Omron Sysmac Studio project medina sin node con todo (Sysmac Studio 1.64.0.64008, StandardProject)

# Controller new_Controller_0: NX102-1020 version 1.60
Axis MC_Axis000, settings changed from default: AxisType=ServoType, FunctionLimit=SingleAxisPTP, UnitsConversion=EnumElement5, UnitsNumerator=8388608, ReducerUse=EnumElement2, TravelDistancePerWorkRotation=180, WorkGearRatio=100, MotorGearRatio=198, MaxVelocity=20, MaxJogVelocity=20, CountMode=EnumElement2, ModuloMAXPosition=360, ModuloMINPosition=0, EncoderTypes=Abs
Axis MC_Axis001, settings changed from default: AxisNumber=1, AxisType=ServoType, FunctionLimit=SingleAxisPTP, UnitsConversion=EnumElement2, UnitsNumerator=8388608, UnitsDenominator=290, MaxVelocity=10, MaxJogVelocity=10, EncoderTypes=Abs
Task PrimaryTask (priority 4, period or condition 2000): Programa0, main
Task PeriodicTask0 (priority 17, period or condition 20000): AMR
Library TMEthernetIP_v2.0.0 2.0.0 (contents left out)
Library ARCL_Comms_Lib 1.3.0 (contents left out)

TYPE RfidCommand : STRUCT
    CommExec : WORD;
    CmdCode : WORD;
    CmdParam1 : WORD;
    CmdParam2 : WORD;
    CmdData : array[0..15] of word;
END_STRUCT END_TYPE
TYPE RfidResponse : STRUCT
    RfidStatus : WORD;
    RfidErrorCode : WORD;
    RfidRespInfo1 : WORD;
    RfidRespInfo2 : WORD;
    RfidRespData : array[0..15] of WORD;
END_STRUCT END_TYPE
TYPE RFID_Status : UNION
    Status_reg : word;
    Status_bits : ARRAY[0..15] OF BOOL;
END_UNION END_TYPE
TYPE CmdRFID : (Read_ID := 1, Read_data := 2, Write_Data := 3, LockRfid := 4, Data_fill := 5, Overwrite_control := 6, Restore_data := 7, Copy_data := 8, Initialize := 4096, Set_RF_Comm_Settings := 4097, Get_RF_tag_comm := 4098, Set_multi_Reades := 4099, Get_multi_reader := 4100, Get_model_information := 8192, Get_firmware_version := 8193, Get_operating_time := 8194, Measure_noise := 8195, Get_comd_error_log := 8196, Get_restore_infomation := 8197, Get_multireader_status := 8198, Reset := 12288); END_TYPE
TYPE Status_struct : STRUCT
    Datos_bits : ARRAY[0..15] OF BOOL;
END_STRUCT END_TYPE
TYPE stCarouselSlot : STRUCT
    RoomID : INT;
    MedID : INT;
    IsLoaded : BOOL;
    IsDelivered : BOOL;
END_STRUCT END_TYPE

VAR_GLOBAL
    DataFromRFID : RfidResponse;  (* network input *)
    ArrayFromTM : array[0..491] of byte;  (* network input *)
    ArrayToTM : array[0..295] of byte;  (* network output *)
    StructFromTM : ATC_E\TMEthernetIP\FromTM;
    StructToTM : ATC_E\TMEthernetIP\ToTM;
    DataToRFID : RfidCommand;  (* network output *)
END_VAR
VAR_GLOBAL CONSTANT
    MC_Axis000 : _sAXIS_REF;  (* at MC://_MC_AX[0] *)
    MC_Axis001 : _sAXIS_REF;  (* at MC://_MC_AX[1] *)
END_VAR
VAR_GLOBAL
    habitaciones : ARRAY[0..9] OF int;  (* network output *)
    medicamentos : ARRAY[0..9] OF int;  (* network output *)
    test_escritura : INT;  (* published *)
    Carrusel : ARRAY[0..9] OF stCarouselSlot;
    etapa : INT;
    activar : BOOL;
    done_amr : BOOL;
    pos_carrusel : LREAL;
    pos_trampilla : LREAL;
    done_carrusel : BOOL;
    done_trampilla : BOOL;
    boton_recogido_HMI : BOOL;
    trampilla : BOOL;
    trampilla1 : BOOL;
    pos_amr : STRING[25];
    NodeRed_StartMission : BOOL;  (* published *)
    NodeRed_listo : BOOL;  (* published *)
    doneRFID : BOOL;
    RFID_RoomID : INT;
    miARCL : ARCL_Comms_Lib\ARCL_ST_Connection;
    MedID_Actual : INT;  (* published *)
    Habitacion_Actual : INT;  (* published *)
    Nombre_Medicamento : STRING[30];  (* published *)
    StartMission_Manual : BOOL;
    Sin_Pedidos : BOOL;
END_VAR

PROGRAM main
VAR
    TM_Done : BOOL;
    PLC_Listo : BOOL;
    fase_reparto : BOOL;
    CurrentSlot : INT;
    TargetRoom : INT;
    i : INT;
    var1 : INT;
    DoctorRFID_ID : INT;
    sub_etapa_carga : INT;
    cargas_realizadas : INT;
    total_cargas_pendientes : INT;
    stock_medicamentos : ARRAY[1..5] OF INT;
END_VAR
VAR_EXTERNAL
    activar : BOOL;
    NodeRed_listo : BOOL;
    habitaciones : ARRAY[0..9] OF int;
    medicamentos : ARRAY[0..9] OF int;
    NodeRed_StartMission : BOOL;
    pos_amr : STRING[25];
    done_amr : BOOL;
    pos_trampilla : LREAL;
    done_trampilla : BOOL;
    etapa : INT;
    pos_carrusel : LREAL;
    Carrusel : ARRAY[0..9] OF stCarouselSlot;
    done_carrusel : BOOL;
    doneRFID : BOOL;
    RFID_RoomID : INT;
    trampilla : BOOL;
    boton_recogido_HMI : BOOL;
    trampilla1 : BOOL;
    StructToTM : ATC_E\TMEthernetIP\ToTM;
    StructFromTM : ATC_E\TMEthernetIP\FromTM;
    DataFromRFID : RfidResponse;
    MedID_Actual : INT;
    Habitacion_Actual : INT;
    Nombre_Medicamento : STRING[30];
    StartMission_Manual : BOOL;
    Sin_Pedidos : BOOL;
END_VAR
// ============================================================================
// MAQUINA DE ESTADOS AMR + CARRUSEL + TM  (adaptada al ladder del proyecto)
// ----------------------------------------------------------------------------
// El ladder mueve los equipos segun el valor de "etapa" (el Execute se mantiene
// a TRUE mientras dura la etapa, con 300 ms de retardo):
//     etapa 10, 60, 100 -> AMR  (ARCL_Goto, destino = pos_amr)       -> done_amr
//     etapa 30, 80      -> Carrusel (servo, destino = pos_carrusel)  -> done_carrusel
//     etapa 20, 40      -> Trampilla (servo, destino = pos_trampilla)-> done_trampilla
//     etapa 25          -> Lector RFID (Rfid01)                      -> doneRFID
//
// Un servo solo hace un movimiento nuevo cuando su Execute pasa de FALSE a TRUE.
// Por eso cada movimiento del carrusel es UNA VISITA NUEVA a la etapa 30 o 80:
// entre un movimiento y el siguiente el programa pasa por una etapa sin motor
// (28 / 32 / 75), el Execute baja y vuelve a subir.
//
// VARIABLES: fase_reparto (BOOL) es LOCAL nueva del programa "main".
// StartMission_Manual y Sin_Pedidos (BOOL) pasan a ser GLOBALES (VAR_EXTERNAL aqui)
// para que la HMI pueda iniciar la mision y mostrar el aviso. El resto ya existia.
//
// Etapas:
//   0 espera orden          10 AMR a Doctor          20 abre trampilla
//  25 RFID (doctor / hab.)  28 elegir ranura         30 mueve carrusel
//  32 espera al doctor      50 elegir entrega        60 AMR a habitacion
//  75 handshake TM          76 espera fin TM         80 carrusel a la ranura
//  90 espera al paciente   100 AMR a base
// ============================================================================

// LA TRAMPILLA SIEMPRE QUEDA ABIERTA:
// posicion fija a 0.0 y nunca se manda cerrar (la etapa 40 no se usa).
pos_trampilla := 0.0;
trampilla := FALSE;
trampilla1 := FALSE;

CASE etapa OF

    // ==========================================
    // 0: ESPERA DE NUEVA ORDEN (MANUAL)
    // ==========================================
    0:
        PLC_Listo := TRUE;
        activar := TRUE;          // alimenta ARCL, servos y comunicacion con el TM
        fase_reparto := FALSE;

        IF StartMission_Manual THEN

            // Contar pedidos validos (habitacion 1..5)
            total_cargas_pendientes := 0;
            FOR i := 0 TO 9 DO
                IF habitaciones[i] >= 1 AND habitaciones[i] <= 5 THEN
                    total_cargas_pendientes := total_cargas_pendientes + 1;
                END_IF;
            END_FOR;

            StartMission_Manual := FALSE;

            IF total_cargas_pendientes = 0 THEN
                Sin_Pedidos := TRUE;          // sin pedidos: no arranca
            ELSE
                Sin_Pedidos := FALSE;
                PLC_Listo := FALSE;

                FOR i := 0 TO 9 DO
                    IF habitaciones[i] >= 1 AND habitaciones[i] <= 5 THEN
                        Carrusel[i].RoomID := habitaciones[i];
                    ELSE
                        Carrusel[i].RoomID := 0;
                    END_IF;
                    Carrusel[i].MedID := medicamentos[i];
                    Carrusel[i].IsLoaded := FALSE;
                    Carrusel[i].IsDelivered := FALSE;
                END_FOR;

                cargas_realizadas := 0;
                CurrentSlot := 0;
                etapa := 10;
            END_IF;
        END_IF;

    // ==========================================
    // FASE DE CARGA EN CONSULTORIO (DOCTOR)
    // ==========================================
    10: // AMR VA AL CONSULTORIO DEL DOCTOR
        pos_amr := 'Doctor';
        IF done_amr THEN
            etapa := 20;
        END_IF;

    20: // ABRIR TRAMPILLA (se queda abierta toda la mision)
        IF done_trampilla THEN
            boton_recogido_HMI := FALSE;
            etapa := 25;
        END_IF;

    25: // RFID: lectura del doctor (fase de carga) o de la puerta (fase de reparto)
        var1 := WORD_TO_INT(In := DataFromRFID.RfidRespData[0]);

        IF NOT fase_reparto THEN
            IF doneRFID OR (var1 <> 0 AND var1 = DoctorRFID_ID) THEN
                CurrentSlot := 0;
                etapa := 28;
            END_IF;
        ELSE
            IF doneRFID OR (var1 <> 0 AND var1 = TargetRoom) THEN
                etapa := 75;
            END_IF;
        END_IF;

    28: // ELEGIR LA SIGUIENTE RANURA QUE HAY QUE CARGAR (sin motores)
        IF CurrentSlot <= 9 THEN
            IF Carrusel[CurrentSlot].RoomID > 0 AND NOT Carrusel[CurrentSlot].IsLoaded THEN

                MedID_Actual := Carrusel[CurrentSlot].MedID;
                Habitacion_Actual := Carrusel[CurrentSlot].RoomID;

                CASE MedID_Actual OF
                    1: Nombre_Medicamento := 'Paracetamol';
                    2: Nombre_Medicamento := 'Ibuprofeno';
                    3: Nombre_Medicamento := 'Antibiotico';
                    4: Nombre_Medicamento := 'Suero';
                    5: Nombre_Medicamento := 'Insulina';
                ELSE
                    Nombre_Medicamento := 'Desconocido';
                END_CASE;

                etapa := 30;
            ELSE
                CurrentSlot := CurrentSlot + 1;
            END_IF;
        ELSE
            // Todas las ranuras cargadas: empieza el reparto (trampilla sigue abierta)
            CurrentSlot := 0;
            fase_reparto := TRUE;
            etapa := 50;
        END_IF;

    30: // CARRUSEL A LA RANURA (el ladder mueve el servo en esta etapa)
        pos_carrusel := CurrentSlot * 36.0;
        IF done_carrusel THEN
            boton_recogido_HMI := FALSE;      // descarta pulsaciones anteriores
            etapa := 32;
        END_IF;

    32: // ESPERA AL DOCTOR (pulsador HMI)
        IF boton_recogido_HMI THEN
            Carrusel[CurrentSlot].IsLoaded := TRUE;
            cargas_realizadas := cargas_realizadas + 1;
            boton_recogido_HMI := FALSE;
            CurrentSlot := CurrentSlot + 1;
            etapa := 28;
        END_IF;

    // ==========================================
    // FASE DE REPARTO MULTI-HABITACION
    // ==========================================
    50: // BUSCAR LA SIGUIENTE ENTREGA PENDIENTE
        TargetRoom := 0;

        FOR i := 0 TO 9 DO
            IF Carrusel[i].IsLoaded AND NOT Carrusel[i].IsDelivered THEN
                TargetRoom := Carrusel[i].RoomID;
                CurrentSlot := i;
                EXIT;
            END_IF;
        END_FOR;

        IF TargetRoom > 0 THEN
            etapa := 60;
        ELSE
            etapa := 100;         // mision completa
        END_IF;

    60: // AMR VIAJA A LA HABITACION
        CASE Carrusel[CurrentSlot].RoomID OF
            1: pos_amr := 'habitacion1';
            2: pos_amr := 'habitacion2';
            3: pos_amr := 'habitacion3';
            4: pos_amr := 'habitacion4';
            5: pos_amr := 'habitacion5';
        END_CASE;

        IF done_amr THEN
            etapa := 25;          // lectura RFID de la puerta (fase_reparto = TRUE)
        END_IF;

    75: // HANDSHAKE ROBOT TM (24 -> 22)
        StructToTM.TM_4_O2T_RegisterInt.O2T_Register_Int[0] := 24;

        IF StructFromTM.TM_9_T2O_RegisterInt.T2O_Register_Int[0] = 22 THEN

            IF Carrusel[CurrentSlot].MedID >= 1 AND Carrusel[CurrentSlot].MedID <= 5 THEN
                IF stock_medicamentos[Carrusel[CurrentSlot].MedID] > 0 THEN
                    stock_medicamentos[Carrusel[CurrentSlot].MedID] := stock_medicamentos[Carrusel[CurrentSlot].MedID] - 1;
                END_IF;
            END_IF;

            StructToTM.TM_4_O2T_RegisterInt.O2T_Register_Int[0] := 0;
            i := 0;
            etapa := 76;
        END_IF;

    76: // ESPERAR A QUE EL TM SUELTE EL 22 (si no, la siguiente entrega se daria por confirmada)
        i := i + 1;
        IF StructFromTM.TM_9_T2O_RegisterInt.T2O_Register_Int[0] <> 22 OR i >= 500 THEN
            etapa := 80;
        END_IF;

    80: // CARRUSEL A LA RANURA DE ESTA ENTREGA (el ladder mueve el servo; trampilla ya abierta)
        pos_carrusel := CurrentSlot * 36.0;
        IF done_carrusel THEN
            boton_recogido_HMI := FALSE;
            etapa := 90;
        END_IF;

    90: // ENTREGA AL PACIENTE (trampilla abierta)
        IF boton_recogido_HMI THEN
            Carrusel[CurrentSlot].IsDelivered := TRUE;
            boton_recogido_HMI := FALSE;
            etapa := 50;          // siguiente entrega
        END_IF;

    // ==========================================
    // FASE DE RETORNO
    // ==========================================
    100: // VOLVER A BASE
        pos_amr := 'base';
        IF done_amr THEN
            etapa := 0;
        END_IF;

END_CASE;
END_PROGRAM

PROGRAM Programa0
VAR
    DatosDelTM_Enalbe : BOOL;
    DatosDelTM_Instancia : ATC_E\TMEthernetIP\ConvertDataFromTM;
    DatosDelTM_Done : BOOL;
    DatosAlTM_Enable : BOOL;
    DatosAlTm_Done : BOOL;
    DatosAlTM_Instancia : ATC_E\TMEthernetIP\ConvertDataToTM;
    Rfid01 : RfidOperation;
    Start_servo_01 : BOOL;
    iPowerServo01 : MC_Power;
    servo1Home : BOOL;
    iServo01HOme : MC_Home;
    servo01Giro : BOOL;
    iServo01Giro : MC_MoveAbsolute;
    noHacer : BOOL;
    ErrorGiro : BOOL;
    ErrorHoming : BOOL;
    ErrorPower : BOOL;
    ErrorIDPower : WORD;
    ErrorIDGiro : WORD;
    consignaPosicion : LREAL;
    iMc_reset : MC_Reset;
    bReset : BOOL;
    iARCLConnect : ARCL_Comms_Lib\ARCL_Connect;
    ipAMR : STRING[20] := '192.168.20.173';
    portAMR : UINT := 7171;
    passAMR : STRING[30] := 'omron';
    connAMR : STRING[10] := 'ld90';
    miARCL : ARCL_Comms_Lib\ARCL_ST_Connection;
    AMR_busy : BOOL;
    AMR_error : BOOL;
    AMR_ErrorID : WORD;
    AMR_Status : STRING[30];
    iAMRGoto : ARCL_Comms_Lib\ARCL_Goto;
    miGoal : STRING[25] := 'PruebaGoal';
    AMRGotoBusy : BOOL;
    AMRGotoError : BOOL;  (* AMRGotoErrorID *)
    AMRGotoID : WORD;
    AMRGotoStatus : STRING[30];
    iPowerServo02 : MC_Power;
    Start_servo_02 : BOOL;
    ErrorPowerServo01 : BOOL;  (* ErrorIDPowerServo01 *)
    bResetServo01 : BOOL;
    servo2Home : BOOL;
    bResetServo02 : BOOL;
    iMC_Reset_02 : MC_Reset;
    iMC_HomeServo02 : MC_Home;
    iMC_MoveAbsolute_02 : MC_MoveAbsolute;
    servo02Giro : BOOL;
    ErrorGiroServo02 : BOOL;
    ErrorIDServo02 : WORD;
    consignaPosicion02 : LREAL;
    noEjecutar : BOOL;
    t1 : TON;
    vel_trampilla : LREAL := 10;
    ace_trampilla : LREAL := 10;
    des_trampilla : LREAL := 10;
    jerk_trampilla : LREAL := 10;
    velocidad_carrusel : LREAL := 20;
    acceleracion_carrusel : LREAL := 10;
    desaceleracion_carrusel : LREAL := 10;
    jerk_carrusel : LREAL := 10;
    temp5 : TON;
    temp4 : TON;
    prueba : BOOL;
    prueb1 : BOOL;
    mc_trampilla : MC_MoveAbsolute;
END_VAR
VAR_EXTERNAL
    ArrayFromTM : array[0..491] of byte;
    StructFromTM : ATC_E\TMEthernetIP\FromTM;
    StructToTM : ATC_E\TMEthernetIP\ToTM;
    ArrayToTM : array[0..295] of byte;
END_VAR
VAR_EXTERNAL CONSTANT
    MC_Axis000 : _sAXIS_REF;
    MC_Axis001 : _sAXIS_REF;
END_VAR
VAR_EXTERNAL
    pos_carrusel : LREAL;
    pos_trampilla : LREAL;
    done_carrusel : BOOL;
    done_trampilla : BOOL;
    activar : BOOL;
    etapa : INT;
    trampilla : BOOL;
    trampilla1 : BOOL;
    doneRFID : BOOL;
    DataToRFID : RfidCommand;
END_VAR

(* Section Servos: ladder, written here as Structured Text *)

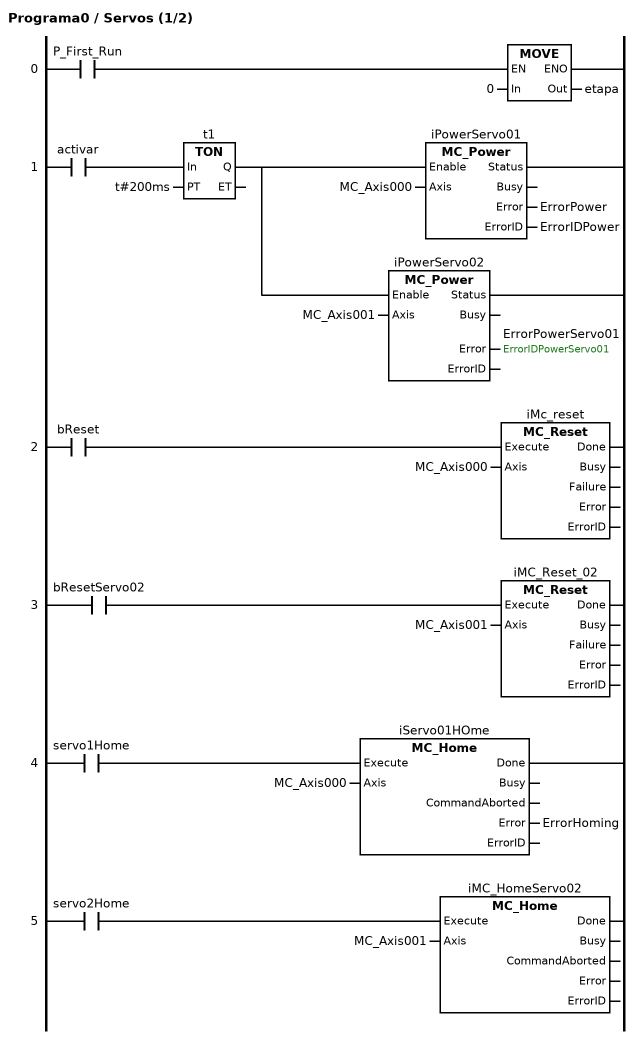
(* Rung 0 *)
IF P_First_Run THEN etapa := 0; END_IF;
(* Rung 1 *)
t1(In := activar, PT := t#200ms);
iPowerServo01(Enable := t1.Q, Axis := MC_Axis000, Error => ErrorPower, ErrorID => ErrorIDPower);
iPowerServo02(Enable := t1.Q, Axis := MC_Axis001, Error => ErrorPowerServo01);
(* Rung 2 *)
iMc_reset(Execute := bReset, Axis := MC_Axis000);
(* Rung 3 *)
iMC_Reset_02(Execute := bResetServo02, Axis := MC_Axis001);
(* Rung 4 *)
iServo01HOme(Execute := servo1Home, Axis := MC_Axis000, Error => ErrorHoming);
(* Rung 5 *)
iMC_HomeServo02(Execute := servo2Home, Axis := MC_Axis001);

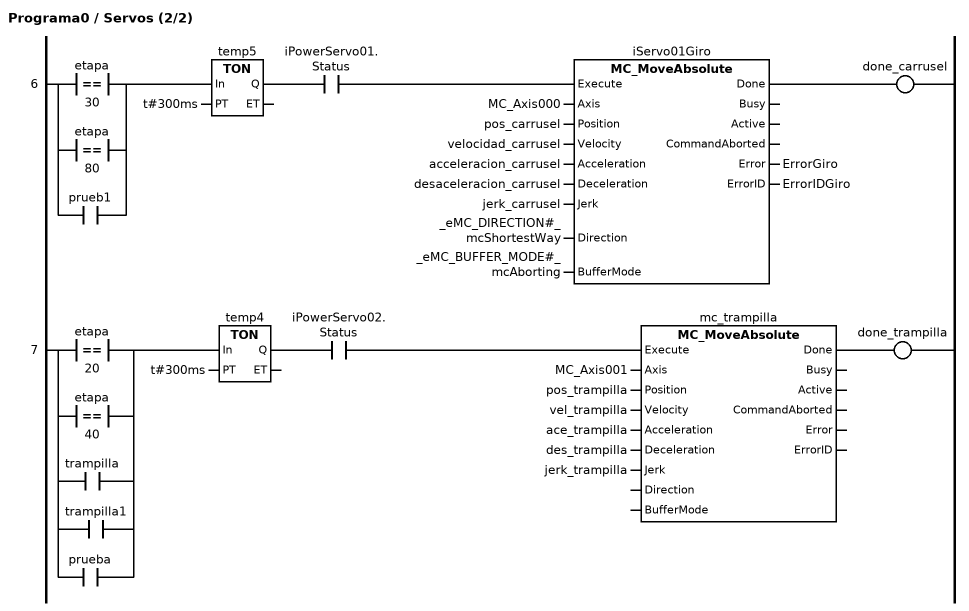
(* Rung 6 *)
temp5(In := (etapa = 30) OR (etapa = 80) OR prueb1, PT := t#300ms);
iServo01Giro(Execute := temp5.Q AND iPowerServo01.Status, Axis := MC_Axis000, Position := pos_carrusel, Velocity := velocidad_carrusel, Acceleration := acceleracion_carrusel, Deceleration := desaceleracion_carrusel, Jerk := jerk_carrusel, Direction := _eMC_DIRECTION#_mcShortestWay, BufferMode := _eMC_BUFFER_MODE#_mcAborting, Error => ErrorGiro, ErrorID => ErrorIDGiro);
done_carrusel := iServo01Giro.Done;
(* Rung 7 *)
temp4(In := (etapa = 20) OR (etapa = 40) OR trampilla OR trampilla1 OR prueba, PT := t#300ms);
mc_trampilla(Execute := temp4.Q AND iPowerServo02.Status, Axis := MC_Axis001, Position := pos_trampilla, Velocity := vel_trampilla, Acceleration := ace_trampilla, Deceleration := des_trampilla, Jerk := jerk_trampilla);
done_trampilla := mc_trampilla.Done;

(* Section RFID: ladder, written here as Structured Text *)

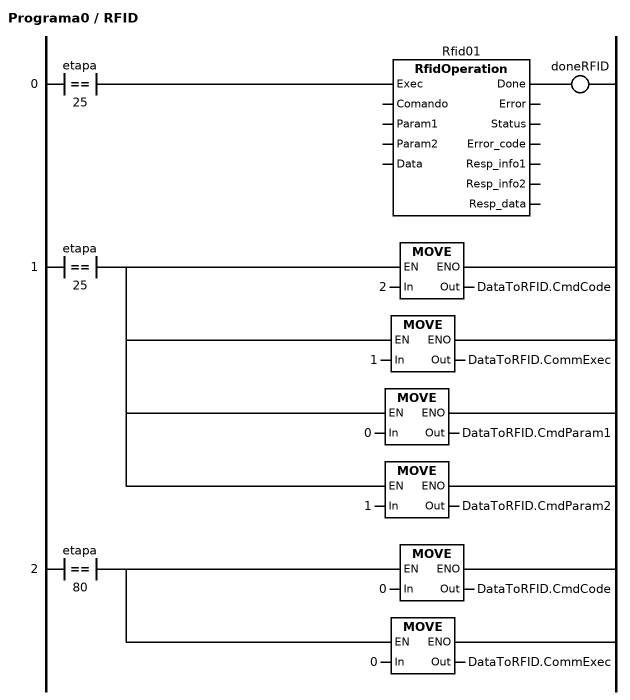
(* Rung 0 *)
Rfid01(Exec := etapa = 25);
doneRFID := Rfid01.Done;
(* Rung 1 *)
IF etapa = 25 THEN
    DataToRFID.CmdCode := 2;
    DataToRFID.CommExec := 1;
    DataToRFID.CmdParam1 := 0;
    DataToRFID.CmdParam2 := 1;
END_IF;
(* Rung 2 *)
IF etapa = 80 THEN
    DataToRFID.CmdCode := 0;
    DataToRFID.CommExec := 0;
END_IF;

(* Section RobotTM: ladder, written here as Structured Text *)

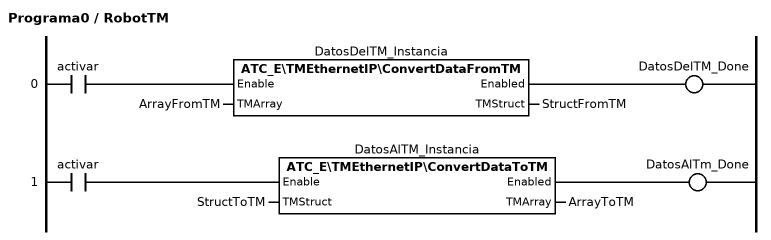
(* Rung 0 *)
DatosDelTM_Instancia(Enable := activar, TMArray := ArrayFromTM, TMStruct => StructFromTM);
DatosDelTM_Done := DatosDelTM_Instancia.Enabled;
(* Rung 1 *)
DatosAlTM_Instancia(Enable := activar, TMStruct := StructToTM, TMArray => ArrayToTM);
DatosAlTm_Done := DatosAlTM_Instancia.Enabled;
END_PROGRAM

PROGRAM AMR
VAR
    CONECTAR : ARCL_Comms_Lib\ARCL_Connect;
    T2 : TON;
    IR_A : ARCL_Comms_Lib\ARCL_Goto;
    T3 : TON;
    ipAMR : STRING[20] := '192.168.20.130';
    portAMR : UINT := 7171;
    passAMR : STRING[30] := 'omron';
    ReconectionTime : TIME := t#5s;
    connAMR : STRING[10] := 'PLC1';
    fast : BOOL;
    timeout : TIME := T#200S;
    heading : INT := 0;
    default : BOOL := True;
END_VAR
VAR_EXTERNAL
    miARCL : ARCL_Comms_Lib\ARCL_ST_Connection;
    activar : BOOL;
    done_amr : BOOL;
    etapa : INT;
    pos_amr : STRING[25];
END_VAR

(* Section LD90: ladder, written here as Structured Text *)

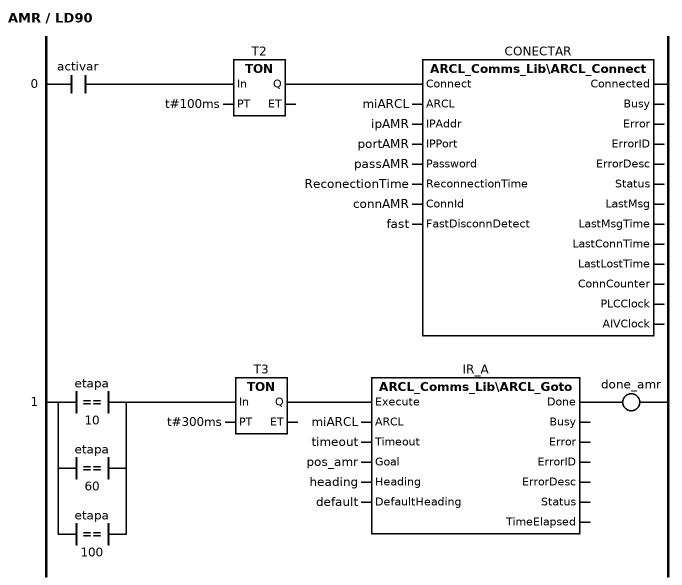
(* Rung 0 *)
T2(In := activar, PT := t#100ms);
CONECTAR(Connect := T2.Q, ARCL := miARCL, IPAddr := ipAMR, IPPort := portAMR, Password := passAMR, ReconnectionTime := ReconectionTime, ConnId := connAMR, FastDisconnDetect := fast);
(* Rung 1 *)
T3(In := (etapa = 10) OR (etapa = 60) OR (etapa = 100), PT := t#300ms);
IR_A(Execute := T3.Q, ARCL := miARCL, Timeout := timeout, Goal := pos_amr, Heading := heading, DefaultHeading := default);
done_amr := IR_A.Done;
END_PROGRAM

FUNCTION_BLOCK RfidOperation
VAR
    estado_RFID : RFID_Status;
    paso : UINT;
END_VAR
VAR_INPUT
    Exec : BOOL;
    Comando : WORD;
    Param1 : WORD;
    Param2 : WORD;
    Data : ARRAY[0..15] OF word;
END_VAR
VAR_OUTPUT
    Done : BOOL;
    Error : BOOL;
    Status : WORD;
    Error_code : WORD;
    Resp_info1 : WORD;
    Resp_info2 : WORD;
    Resp_data : ARRAY[0..15] OF word;
END_VAR
VAR_EXTERNAL
    DataFromRFID : RfidResponse;
    DataToRFID : RfidCommand;
END_VAR
// 0. ACTUALIZACIÓN DE LA UNIÓN INTERNA
// Sincronizamos la palabra de estado recibida por red con nuestra unión para procesar bits
estado_RFID.Status_reg := DataFromRFID.RfidStatus;

CASE Paso OF
    0: // --- ESPERA DE ORDEN ---
        // Comprobamos que el lector esté READY (Bit 0) y no BUSY (Bit 1)
        IF estado_RFID.Status_bits[0] AND NOT estado_RFID.Status_bits[1] AND Exec THEN
            // 1. Cargamos comando y parámetros en la estructura de salida global
            DataToRFID.CmdCode   := Comando;
            DataToRFID.CmdParam1 := Param1;
            DataToRFID.CmdParam2 := Param2;
            
            // Si el comando es de escritura (3), copiamos el array de datos
            IF Comando = 16#0003 THEN
                DataToRFID.CmdData := Data; 
            END_IF;

            // 2. Activamos el bit EXE (Bit 0 de CommExec)
            // Asignamos 1 al Word para poner el Bit 0 a TRUE
            DataToRFID.CommExec := 16#0001; 
            
            // Limpiamos salidas de estado del FB
            Done  := FALSE;
            Error := FALSE;
            Paso  := 10;
        END_IF;

    10: // --- ESPERA DE CONFIRMACIÓN (BUSY) ---
        // El lector indica que ha recibido la orden activando BUSY (Bit 1)
        IF estado_RFID.Status_bits[1] THEN
            Paso := 20;
        END_IF;

    20: // --- PROCESAMIENTO Y RESULTADO ---
        // Esperamos a que finalice: NORM (Bit 2) o ERR (Bit 3)
        IF estado_RFID.Status_bits[2] OR estado_RFID.Status_bits[3] THEN
            
            // Mapeamos los resultados a tus salidas del FB
            Status     := estado_RFID.Status_reg;
            Error_code := DataFromRFID.RfidErrorCode;
            Resp_info1 := DataFromRFID.RfidRespInfo1;
            Resp_info2 := DataFromRFID.RfidRespInfo2;

            // Si terminó con éxito (NORM), capturamos los datos leídos
            IF estado_RFID.Status_bits[2] THEN
                Resp_data := DataFromRFID.RfidRespData;
                Done      := TRUE;
            END_IF;

            // Si terminó con error (ERR)
            IF estado_RFID.Status_bits[3] THEN
                Error := TRUE;
            END_IF;

            // 3. Cierre del Handshake: Bajamos el bit EXE
            DataToRFID.CommExec := 16#0000;
            Paso := 30;
        END_IF;

    30: // --- FINALIZACIÓN Y REARME ---
        // Esperamos a que el lector limpie el estado y vuelva a READY
        IF estado_RFID.Status_bits[0] AND NOT estado_RFID.Status_bits[1] THEN
            // Solo permitimos reiniciar si el usuario ha bajado la entrada 'Exec'
            IF NOT Exec THEN
                Done := FALSE;
                Paso := 0;
            END_IF;
        END_IF;
END_CASE;
END_FUNCTION_BLOCK

# Device HMI_NA5_1 (NA): not converted